PROGRAM main
  VAR
    Button AT %QX0.0 : BOOL;
    Motor AT %QX0.1 : BOOL;
    Package_sense AT %QX0.2 : BOOL;
    reset_counter AT %QX0.3 : BOOL;
    total_count AT %MW1 : INT;
    Bigboxcount AT %MW2 : INT;
    Mediumboxcount AT %MW3 : INT;
    Smallboxcount AT %MW4 : INT;
    Weight_sensor AT %MW0 : INT;
    CTU0 : CTU;
    CTU1 : CTU;
    is_big AT %MX0.0 : BOOL;
    is_small AT %IXNaN.1 : BOOL;
  END_VAR
  VAR  (* added by the conversion: wires and edge detectors of the diagram *)
    _ADD22_OUT : ANY;
  END_VAR

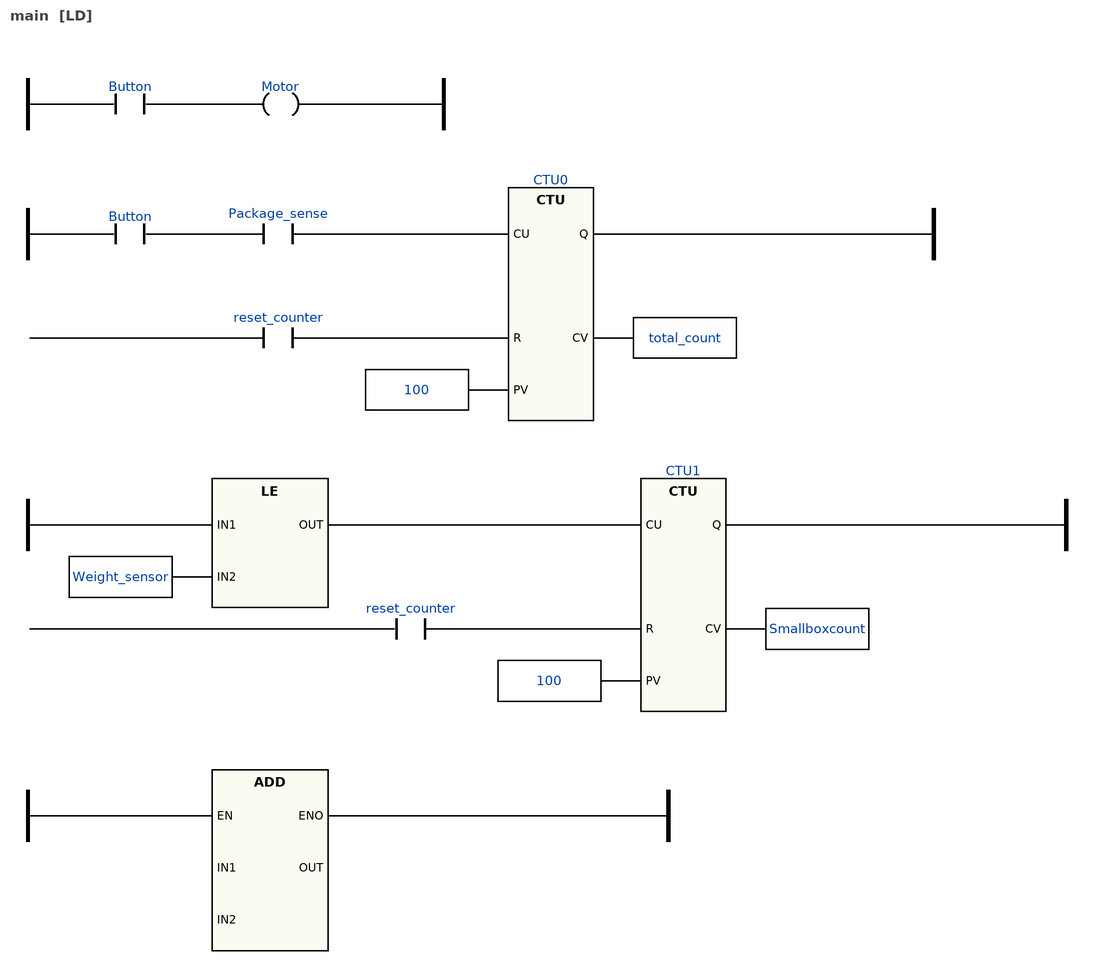
(* LD diagram, written out as Structured Text *)
Motor := Button;
CTU0(CU := Button AND Package_sense, R := reset_counter, PV := 100);
total_count := CTU0.CV;
CTU1(CU := TRUE <= Weight_sensor, R := reset_counter, PV := 100);
Smallboxcount := CTU1.CV;
_ADD22_OUT := ADD();
END_PROGRAM
